{attribute 'qualified_only'}
{attribute 'strict'}
{attribute 'to_string'}
TYPE EN_Pump_SPAL_Operating_Status :
(
	Normal,
	Derated,
	Not_Operable,
	Not_Available
);
END_TYPE

(* stored: Version 1.1.0.1
   DUT EN_Pump_SPAL_Operating_Status: Id {5698ca33-11ec-4565-a0e2-3948daf1d43e} *)
